Staubli VAL3: robotStatus.dtx

public bool _bHeavyAlarm
public bool bAlarmAck
public bool bGOTO
public bool bInSwitch
public bool bIsCycle
public bool bIsError
public bool bIsEstop
public bool bIsHome
public bool bIsMoving
public bool bIsPause
public bool bIsReady
public bool bIsRemoteAuto
public bool bIsSaving
public bool bPowerON
public bool bProgGOTO
public bool bQuitApp
public bool bReloadIO
public bool bSimulate
public bool bToPause
public bool bToStartCycle
public bool bToStopCycle
public num _nAlarmCode[10] = 300
num _nAlarmIndex
public num _nAvgCapacity
public num _nBestCapacity
public num _nCTIndex
public num _nCapacity
public num _nCycleTime
public num _nErrIndex[10]
  [1] = -1
  [2] = -1
  [3] = -1
  [4] = -1
  [5] = -1
  [6] = -1
  [7] = -1
  [8] = -1
  [9] = -1
public num _nOmacStat = 9
public num nActCode
public num nCycleCmd
public num nCycleIndex = 78
public num nCycleMoveID
public num nFrameIndex
public num nHMIcmd
public num nHWState
public num nHeavyAlarmLev
public num nPLCcmd
public num nProgCode = 4
public num nProgFb = 1
public num nSetSwitchValue
public num nToolIndex
public num nTrajCode
public string _sRobotStatus = "错误：-300. :0traj数据库加载错误"
public string sAlarmMes[10]
public string sBusUsing = "PROFINET"
public string sCycleItem = "04 sls"
public string sIOStatus
string sLstIOStatus
string sLstRobStatus
string sLstTrajStatus
public string sPageUsing
public string sTrajStatus = "[04 sls]移动到:78, DOUT[11]-喷涂完成=FALSE"
